           #statBlk := BLKMOV(SRCBLK := #identData, DSTBLK => #statWriteData);
           //Fill with data
           #statDat[4] := #statWriteData[#statWriteOffset];
           #statDat[5] := #statWriteData[1 + #statWriteOffset];
           #statDat[6] := #statWriteData[2 + #statWriteOffset];
           #statDat[7] := #statWriteData[3 + #statWriteOffset];
           #statDat[8] := #statWriteData[4 + #statWriteOffset];
           #statDat[9] := #statWriteData[5 + #statWriteOffset];
           #statDat[10] := #statWriteData[6 + #statWriteOffset];
           #statDat[11] := #statWriteData[7 + #statWriteOffset];
           #statDat[12] := #statWriteData[8 + #statWriteOffset];
           #statDat[13] := #statWriteData[9 + #statWriteOffset];
           #statDat[14] := #statWriteData[10 + #statWriteOffset];
           #statDat[15] := #statWriteData[11 + #statWriteOffset];
           #statDat[16] := #statWriteData[12 + #statWriteOffset];
           #statDat[17] := #statWriteData[13 + #statWriteOffset];
           #statDat[18] := #statWriteData[14 + #statWriteOffset];
           #statDat[19] := #statWriteData[15 + #statWriteOffset];
           #statDat[20] := #statWriteData[16 + #statWriteOffset];
           #statDat[21] := #statWriteData[17 + #statWriteOffset];
           #statDat[22] := #statWriteData[18 + #statWriteOffset];
           #statDat[23] := #statWriteData[19 + #statWriteOffset];
           #statDat[24] := #statWriteData[20 + #statWriteOffset];
           #statDat[25] := #statWriteData[21 + #statWriteOffset];
           #statDat[26] := #statWriteData[22 + #statWriteOffset];
           #statDat[27] := #statWriteData[23 + #statWriteOffset];
           #statDat[28] := #statWriteData[24 + #statWriteOffset];
           #statDat[29] := #statWriteData[25 + #statWriteOffset];
           #statDat[30] := #statWriteData[26 + #statWriteOffset];
           #statDat[31] := #statWriteData[27 + #statWriteOffset];

           //#statIOsizeNetto Bytes are reserved for every transfer
       END_IF;
       IF #statBlk = 0 THEN
           #statNState := #statTelegramState;                           //Telegram: Edit the read data
       END_IF;


       //-----------------------------------------------Telegram state----------------------------------------//
       //---------------------------------------------edit received data--------------------------------------//
       //-----------------------------------------------------------------------------------------------------//  

   1: //Telegram    
       IF #statLength > #statIOsizeNetto -1 THEN                 //Only when length of data > 0 can continue  
           IF #statStatusBits[6] THEN                            //IF RFID error has occured
               #tempStatusWord[1] := #statRecDat[1];          //error_RFID
               #tempStatusWord[0] := 16#0011;                          //Error identifier for RFID errors
               #status := #tempStatus;
               #statNState := #statErrorState;
           END_IF;

           //-------------------------- read command is ready------------------------------------------------//

           IF #statStatusBits[7] AND #statStatusBits[0] THEN
               IF #statRecDat[2] = #statAddrWrite[0] AND #statRecDat[3] = #statAddrWrite[1] THEN //received ADR must be ==sent ADR
                   IF #statBlk = 0 THEN
                       IF #statStatusBits[7] AND NOT #statStatusBits[6] THEN
                           #statLength := #statLength - #statIOsizeNetto;
                           //if len is not dividable with #statIOsizeNetto the adr offset has to be changed that the last (length < #statIOsizeNetto) command is done right
                           IF #statDiffToIOsizeNetto <> 0 AND #statLength < #statIOsizeNetto THEN
                               #statByteMove := #statIOsizeNetto - #statDiffToIOsizeNetto;
                           END_IF;
                           #statWriteOffset := #statWriteOffset + #statIOsizeNetto;                                   //offset must be changed
                           #statAddr := INT_TO_WORD(WORD_TO_INT(#statAddr) + #statIOsizeNetto);     //Change the ADR (#statIOsizeNetto Bytes)       
                           #statNState := #statWriteState;                      //Start a new read command
                       ELSE
                           #statNState := #statIdleState;
                       END_IF;
                   ELSE
                       #tempStatusWord[1] := INT_TO_WORD(#statBlk);                 //Error has to BLKMOV occured
                       #tempStatusWord[0] := 16#0001;                           //functions-Error identifier
                       #status := #tempStatus;
                       #statNState := #statErrorState;
                   END_IF;
               END_IF;
           END_IF;

       ELSE
           #statNState := #statIdleState;
           #statBusy := FALSE;
           #statDone := TRUE;
           #done := TRUE;
           #busy := FALSE;

           #statDat[0] := 16#0;                                          //Reset write command
           #InstSetIoPart(ID      := #hwID,
                          OFFSET  := #statAddrOffset,
                          LEN     := #statIOsize,
                          STATUS  => #statIoPartStatus,
                          ERROR   => #statIoPartError,
                          OUTPUTS := #statDat);

       END_IF;
       #InstSetIoPart(ID := #hwID,                              //read data from process image
                      OFFSET := #statAddrOffset,
                      LEN := #statIOsize,
                      STATUS => #statIoPartStatus,
                      ERROR => #statIoPartError,
                      OUTPUTS := #statDat);

       //------------------------------------------------------------------------------------------------------------//
       //-------------------------------------------------Error state------------------------------------------------//
       //---------------------------------------------error has occured----------------------------------------------//

   3://#Error_state
       #tempError := true;
       #error := #tempError;
       #statBusy := false;
       #statTImerIn := false;
       #statNState := #statIdleState;
       #statDone := false;

       #statDat[0] := 16#0;                                          //Reset write command
       #InstSetIoPart(ID      := #hwID,                              
                      OFFSET  := #statAddrOffset,
                      LEN     := #statIOsize,
                      STATUS  => #statIoPartStatus,
                      ERROR   => #statIoPartError,
                      OUTPUTS := #statDat);

   END_CASE;

   //------------------------------------------------------------------------------------------------------------//
   //-------------------------------------------------Timer------------------------------------------------------//
   //------------------------------------------------------------------------------------------------------------//

   #instTon(IN := #statTImerIn,
            PT := #statTimerPT);

   IF #instTon.Q THEN                      //error has occured. No tag on field during the 5 sec.
       #tempStatusWord[1] := 16#8101;                              //tag has left the field
       #tempStatusWord[0] := 16#0001;                              //identifier rfid errors
       #status:=#tempStatus;
       #statNState := #statErrorState;
   END_IF;
END_FUNCTION_BLOCK

FUNCTION_BLOCK "LIOLink_RF200_SwitchAntenna"   // FB4, SCL
TITLE = LRfidIOL_ANT
{ S7_Optimized_Access := 'FALSE' }
FAMILY : S7-300
VERSION : 3.1
// Set Antenna
// IO-Link V1.1
   VAR_INPUT
      execute : Bool;   // start process
      antennaState : Bool;   // set/reset antenna bit
      hwID : Word;   // Hardware identifier
      portAddr : Int;   // Start address of port
      "version" : Int := 11;
   END_VAR
   VAR_OUTPUT
      done : Bool;   // Ready
      busy : Bool;   // Block active
      error : Bool;   // Error has occured
      status : DWord;   // error status
      statusWord AT status : Array[0..1] of Word;
      presence : Bool;
   END_VAR
   VAR
      statExecuteReq : Bool;   // positive edge og execute
      statAntByte : Byte;   // Byte 0, Status byte
      statAntBit AT statAntByte : Array[0..7] of Bool;
      statNState : Int;   // current state
      statLastState : Int;   // last state
      statAntennaOn : Int := 1;   // On state
      statAntennaOff : Int := 2;   // OFF state
      statReadyState : Int := 3;
      statAnt : Array[0..31] of Byte;   // received buffer
      statAddrOffset : Int;   // step for FOR
      statSent : Array[0..31] of Byte;   // sent buffer
      statPresenceBit : Bool;
      statBusy : Bool;
      InstSetIoPart : SETIO_PART;
      statIoPartError : Bool;
      statIoPartStatus : DWord;
      InstGetIoPart : GETIO_PART;
      statIOsize : Int;
   END_VAR
   VAR_TEMP
      tempDone : Bool;
      tempError : Bool;
      tempStatus : DWord;
      tempStatus_W AT tempStatus : Array[0..1] of Word;
   END_VAR
   VAR CONSTANT
      IOL_V10 : Int := 8;
      IOL_V11 : Int := 32;
      VERSION_10 : Int := 10;   // Identifier IO-Link version 1.0
      VERSION_11 : Int := 11;   // Identifier IO-Link version 1.1
   END_VAR
BEGIN
   REGION BLOCK INFO HEADER
       //===============================================================================
       // Siemens / (c)Copyright 2020
       //-------------------------------------------------------------------------------
       // Title:            LIOLink_RF200_SwitchAntenna
       // Function:         Switches the antenna on/off of SIMATIC RF200 readers via IO-Link
       // Library:          LIOLink
       // Author:           Siemens Industry Online Support
       // Tested with:      CPU 317-2 PN/DP FW 3.2
       // Engineering:      TIA Portal V16
       // Restrictions:     --
       // Requirements:     --
       //-------------------------------------------------------------------------------
       // Change log table:
       // Version  | Date       | Expert in charge       | Changes applied
       //----------|------------|------------------------|------------------------------
       // 01.00.00 | 01.07.2013 | Online Support         | First release
       // 01.01.00 | 01.12.2016 | Online Support         | Upgrade to TIA Portal V14
       // 02.00.00 | 01.09.2017 | Online Support         | Upgrade to TIA Portal V14 SP1
       //                                                | Implementation of Programming styleguide
       //                                                | Added support for IO-Link V1.1 readers
       // 02.01.00 | 01.12.2017 | Online Support         | Bug fixes and performance improvements
       // 02.02.00 | 01.03.2020 | Online Support         | Upgrade to TIA Portal V16
       // 02.03.00 | 08.03.2020 | Online Support         | Added input "version" for IO-Link version
       //===============================================================================
   END_REGION

   IF #version = #VERSION_11 THEN                           //determine IO-Link reader version (1.0/1.1) to set offset
       #statIOsize := #IOL_V11;
   ELSE
       #statIOsize := #IOL_V10;
   END_IF;

   #statAddrOffset:=#portAddr;                              //start adress of port
   #InstGetIoPart(ID := #hwID,                              //read data from process image
                  OFFSET := #statAddrOffset,
                  LEN := #statIOsize,
                  STATUS => #statIoPartStatus,
                  ERROR => #statIoPartError,
                  INPUTS := #statAnt);

   #statAntByte:=#statAnt[0];                              //status byte
   #statPresenceBit := #statAntBit[5];                     //Presence bit. Transponder on field
   #presence := #statPresenceBit;
   #busy := #statBusy;

   //------------------------------------If error byte<>0--------------------------------------------------//
   //------------------------------------save the rfid error-----------------------------------------------//

   IF #statAnt[1]<>0 AND #statBusy THEN
     #statAntByte:=#statAnt[1];  
      #statusWord[1]:=BYTE_TO_WORD(#statAntByte);    //error_BLK
      #statusWord[0]:=16#0011;                    //identifier rfid errors
      #statBusy:=false;
      #done:=false;
      #error:=TRUE;
      #statNState:=0;
   END_IF;

   IF NOT #execute THEN
       #done := false;
       #error := false;
       #status := 0;
   END_IF;

   IF #execute AND #execute<>#statExecuteReq THEN //Positive Edge for antenna on
     #statLastState:=0;
     #statBusy:=TRUE;                              //Block active
     #done:=FALSE;                             //reset all output parameters
     #error:=FALSE;
     #status:=0;
     IF #antennaState THEN                          //if antenna then activate the ANTENNA_ON process
       #statNState:=#statAntennaOn;
     ELSIF NOT #antennaState THEN                   //if not antenna then activate the ANTENNA_OFF process 
       #statNState:=#statAntennaOff;
     END_IF;

   END_IF;
   #statExecuteReq:=#execute;


   //---------------------------------------Antenna on state-----------------------------------------------//
   //---------------------------------------Reset Antenna bit----------------------------------------------//

   CASE #statNState OF
       0:  //Idle
           ;
       1:  //Antenna_on
                                                        //Antenna on process
           #statAntBit[4] := false;                        //Reset Byte 0, bit 4
           #statSent[0] := 16#0;
           #statLastState := #statAntennaOn;
           #InstSetIoPart(ID := #hwID,                         //Write data into process image
                          OFFSET := #statAddrOffset,
                          LEN := #statIOsize,
                          STATUS => #statIoPartStatus,
                          ERROR => #statIoPartError,
                          OUTPUTS := #statSent);
           IF NOT #statIoPartError AND #statAnt[1] = 0 THEN
               #statNState := #statReadyState;
           ELSIF #statIoPartError THEN
               #tempError := true;
               #error := #tempError;                             //error has occured
               #statBusy := FALSE;
               #tempStatus_W[1] := DWORD_TO_WORD(#statIoPartStatus);//error_BLK
               #tempStatus_W[0] := 16#0001;                    //identifier block errors
           END_IF;
       2:
                                                      //Antenna off process
           #statAntBit[4] := true;                         //set Byte 0, bit 4
           #statSent[0] := 16#10;
           #statLastState := #statAntennaOff;
           #InstSetIoPart(ID := #hwID,                         //Write data into process image
                          OFFSET := #statAddrOffset,
                          LEN := #statIOsize,
                          STATUS => #statIoPartStatus,
                          ERROR => #statIoPartError,
                          OUTPUTS := #statSent);
           IF NOT #statIoPartError AND #statAnt[1] = 0 THEN
               IF #statAntByte = 16#10 THEN                    //if status_byte=16#10 then antenna off
                   #statNState := #statReadyState;
               END_IF;
           ELSIF #statIoPartError THEN
               #tempError := true;
               #error := #tempError;                              //Error has occured
               #statBusy := FALSE;
               #tempStatus_W[1] := DWORD_TO_WORD(#statIoPartStatus);//error_BLK
               #tempStatus_W[0] := 16#0001;                     //identifier block errors
           END_IF;
       3:
           #tempDone := true;
           #done := #tempDone;                           //Ready
           #statBusy := FALSE;
           #statNState := 0;
   END_CASE;
END_FUNCTION_BLOCK

// folder: LIOLink/S7-1200/1500/Base blocks

FUNCTION_BLOCK "LIOLink_Diagnose"   // FB3, SCL
TITLE = LIOLink_Diagnose
{ S7_Optimized_Access := 'TRUE' }
AUTHOR : SIOS
FAMILY : LIOLink
VERSION : 0.1
// LIOLink_Diagnose is used to read the diagnose of all the ports of any IO-Link-Master Product of Siemens.
   VAR_INPUT
      execute : Bool;   // Rising edge starts the execution of the action once
      hwID : HW_IO;   // Hardware identifier of IO-Link master module or first sub module
      cap : Int;   // Client Access Point (CAP) 0xB400 or 0x00E3 (227)
   END_VAR
   VAR_OUTPUT
      done : Bool;   // TRUE: FB processing successfully completed
      busy : Bool;   // TRUE: FB is active and new output values can be expected.
      error : Bool;   // FALSE: No error / TRUE: An error occurred during the execution of the FB.
      status : Word := 16#7000;   // 16#0000-16#7FFF: Status of the FB / 16#8000-16#FFFF: Error identification (see following table)
      diagnostics : "LIOLink_typeDiagnostics";   // Diagnostics information of FB
      events : "LIOLink_typeEvents";
   END_VAR
   VAR
      statExecuteOld : Bool;   // Previous value of input `execute` for edge detection
      statDone : Bool;   // Static value for output 'done'
      statBusy : Bool;   // Static value for output 'busy'
      statError : Bool;   // Static value for output 'error'
      statStatus : Word;   // Static value for output 'status'
      statSubFunctionStatus : DWord;   // Static value for output 'subFunctionStatus'.
      statFBState : DInt;   // State of the state machine
      statFBErrorState : DInt;   // State in the state machine of the block where the error occurred / Zustand in der Zustandsmaschine des Blocks, in dem der Fehler aufgetreten ist
      statHwID : HW_ANY;   // Static value for input 'HwID'
      statHwIDprevious : HW_IO;   // Static value for input 'hwID' from the previous execute / Statischer Wert für Eingang 'hwID'
      statEmptyDiagnostics : "LIOLink_typeDiagnostics";   // Empty diagnostics information (for initialization purposes only)
      instRdRec : RDREC;   // System function "read data record"
      instRdDiag : RDREC;   // System function "read data record"
      statDiagRecord : Array[0..#LAST_INDEX_DIAG_RECORD] of Byte;   // Data record of port diagnose
      statDiagRecordEco : "LIOLink_typeEvents";
      statCap : UInt;   // Static value for input 'cap'
      statRead : Array[0..231] of Byte;   // Data record, Output of RDREC
      statIndexDiag : UInt;   // Static value for index of data record of port diagnose
      statPortNumber : Int := 8;   // Number of Ports of IO-Link-Master
      statPortEco : UInt := 1;   // Static value for a port counter of EcoPN
   END_VAR
   VAR_TEMP
      tempExecute : Bool;   // Temporary value for input 'execute'
      tempHwID : HW_IO;   // Temporary value for input 'hwID'
      tempCap : Int;   // Temporary value for input 'cap'
      tempPortNumber : Int;   // Temporary value for port number
      tempEventNumber : Int;   // Temporary value for event number
      tempIndexDiagRec : Int;   // Temporary value for index of data record (array) of diagnose
   END_VAR
   VAR CONSTANT
      INDEX_CAP_IOLINK : Word := 16#B000;   // Index of the data record for IOLM_Info. Only IO-Link-Masters with CAP=16#B000 support this call.
      INDEX_DIAG_OTHER : Word := 16#00E5;   // Index for port status based on Siemens Standard (old): 229 => reads status of all ports
      INDEX_DIAG_ECO : Word := 16#B200;   // Index for port status based on IO-Link-Standard: 16#B20n, n:Port number => reads port status of only one port
      CAP_LEGACY : Word := 16#00E3;   // Siemens (old) Standard CAP: 227
      CAP_STANDARD : Word := 16#B400;   // IO-Link Standard CAP: 16#B400
      STATUS_EXECUTION_FINISHED_NO_ERROR : Word := 16#0000;   // Processing finished without error
      STATUS_NO_CALL : Word := 16#7000;   // No current processing request / no order in process
      STATUS_FIRST_CALL : Word := 16#7001;   // First call after new incoming job request (rising edge at 'execute')
      STATUS_SUBSEQUENT_CALL : Word := 16#7002;   // Subfunction call in progress without further detailing
      STATUS_MASK : DWord := 16#00FF_FF00;   // Mask to filter error codes
      STATUS_RESOURCE_BUSY : DWord := 16#0080_C200;   // Status from WRREC/RDREC: Resource is busy
      ERR_UNDEFINED_STATE : Word := 16#8600;   // Error in function due to an undefined state in the state machine
      ERR_RDREC : Word := 16#8602;   // Error: RDREC encountered an error, see "diagnostics"
      FB_STATE_NO_PROCESSING : DInt := 0;   // FB state: No processing
      FB_STATE_READ_CAP : DInt := 1;   // FB state: Read CAP
      FB_STATE_READ_DIAG : DInt := 2;   // FB state: Read diagnose
      MIN_PORT : Int := 1;   // Minimum number of ports
      MAX_PORT : Int := 8;   // Maximum number of ports
      MIN_EVENTS : Int;   // Minimum number of events
      MAX_EVENTS : Int := 4;   // Maximum number of events
      MASTER_PORT_STATUS_V2 : Byte := 16#02;   // Master port status version 2
      MASTER_PORT_STATUS_V3 : Byte := 16#03;   // Master port status version 3
      MASTER_PORT_STATUS_V4 : Byte := 16#04;   // Master port status version 4
      START_INDEX_MASTER_PORT_STATUS_V2 : Int := 28;   // Start index of relevant data in the case of port status version 2
      START_INDEX_MASTER_PORT_STATUS_V3 : Int := 34;   // Start index of relevant data in the case of port status version 3
      START_INDEX_MASTER_PORT_STATUS_V4 : Int := 42;   // Start index of relevant data in the case of port status version 4
      START_INDEX_MASTER_PORT_STATUS_STANDARD : Int := 18;   // Start index of relevant data in case of a IO-Link Standard data record for port status
      START_INDEX_DIAG_RECORD : Int := 0;   // Start index of diagnose record array
      LAST_INDEX_DIAG_RECORD : Int := 231;   // Last index of diagnose record array
      RESET_WORD : Word := 16#0000;   // Reset event codes
      RESET_BYTE : Byte := 16#00;   // Reset byte for statDiagRecord
      STATUS_RDREC_VALID : Byte := 16#00;   // Status Code of RDREC in cased of no error occurs
      BITMASK_ERR_RDREC_B3 : Byte := 16#DE;   // Status Code of RDREC in case of an error when reading a data record
      BITMASK_ERR_RDREC_B2 : Byte := 16#80;   // Status Code of RDREC in case of an error when reading a data record - Error according to IEC 61158-6
      BITMASK_ERR_RDREC_B1 : Byte := 16#B0;   // Status Code of RDREC in case of an error when reading a data record - invalid index (cap)
   END_VAR
BEGIN
   REGION BLOCK INFO HEADER
       //===============================================================================
       // Siemens / (c)Copyright 2023
       //-------------------------------------------------------------------------------
       // Title:            LIOLink_Diagnosis
       // Function:         Reads diagnose of ports of IO-Link-Masters in IO-Link Standard
       // Library:          LIOLink
       // Author:           SUP SPH
       // Tested with:      CPU 1511F-1 PN FW 2.8
       // Engineering:      TIA Portal V16
       // Restrictions:     S7-1200/1500
       // Requirements:     --
       //-------------------------------------------------------------------------------
       // Change log table:
       // Version  | Date       | Expert in charge       | Changes applied
       //----------|------------|------------------------|------------------------------
       // 01.00.00 | 28.02.2023 | SUP SPH                | First release for TIA Portal V16
       // 
       //===============================================================================
   END_REGION


   REGION TRIGGERING
       #tempExecute := #execute; // Work with temporary value / create process image

       IF (#tempExecute = TRUE) AND (#statExecuteOld = FALSE) // Check if FB is triggered
           // FB shall finish current job before new job can be started with rising edge of execute
           AND (#statStatus = #STATUS_NO_CALL)
       THEN
           REGION Initialize data
               // First call; initialize FB
               #statDone := FALSE;
               #statBusy := TRUE;
               #statError := FALSE;
               #statStatus := #STATUS_FIRST_CALL;
               #statSubFunctionStatus := #STATUS_EXECUTION_FINISHED_NO_ERROR;
               #statFBErrorState := 0;
               #diagnostics := #statEmptyDiagnostics;
               //save the hwID from the previous execute
               #statHwIDprevious := #statHwID;

               //reset static variables of Diagnose Records
               FOR #tempPortNumber := #MIN_PORT TO #MAX_PORT DO
                   FOR #tempEventNumber := #MIN_EVENTS TO #MAX_EVENTS DO
                       #statDiagRecordEco."port"[#tempPortNumber].event[#tempEventNumber].eventQualifier.instance := #RESET_BYTE;
                       #statDiagRecordEco."port"[#tempPortNumber].event[#tempEventNumber].eventQualifier.source := FALSE;
                       #statDiagRecordEco."port"[#tempPortNumber].event[#tempEventNumber].eventQualifier.type := #RESET_BYTE;
                       #statDiagRecordEco."port"[#tempPortNumber].event[#tempEventNumber].eventQualifier.mode := #RESET_BYTE;
                       #statDiagRecordEco."port"[#tempPortNumber].event[#tempEventNumber].eventCode := #RESET_WORD;
                   END_FOR;
               END_FOR;
               FOR #tempIndexDiagRec := #START_INDEX_DIAG_RECORD TO #LAST_INDEX_DIAG_RECORD DO
                   #statDiagRecord[#tempIndexDiagRec] := #RESET_BYTE;
               END_FOR;
           END_REGION

           REGION Save inputs
               //save input parameters
               #tempHwID := #hwID;
               #tempCap := #cap;
           END_REGION

           REGION Check parameters
               IF #statStatus = #STATUS_FIRST_CALL THEN // Parameters OK
                   IF #tempCap <> 0 THEN   //check if cap is predefined, or given by the user
                       #statCap := INT_TO_UINT(#tempCap);
                       #statFBState := #FB_STATE_READ_DIAG;
                   ELSIF (#statCap <> WORD_TO_UINT(#CAP_STANDARD) AND #statCap <> WORD_TO_UINT(#CAP_LEGACY)) OR (#statHwIDprevious <> #tempHwID) THEN
                       #statFBState := #FB_STATE_READ_CAP;
                   ELSE //CAP already known
                       #statFBState := #FB_STATE_READ_DIAG;
                   END_IF;
               END_IF;
               //save current hwID
               #statHwID := #tempHwID;
           END_REGION

       ELSIF (#statStatus = #STATUS_FIRST_CALL) THEN
           #statStatus := #STATUS_SUBSEQUENT_CALL;
       ELSIF (#statFBState=#FB_STATE_NO_PROCESSING) THEN
           #statStatus := #STATUS_NO_CALL;
           #statDone := FALSE;
           #statBusy := FALSE;
           #statError := FALSE;

           #instRdDiag(REQ := FALSE,
                       RECORD := #statDiagRecord);

           #instRdRec(REQ := FALSE,
                      RECORD := #statRead);
       END_IF;

       // Edge detection 'execute' input
       #statExecuteOld := #tempExecute;
   END_REGION TRIGGERING

   REGION STATE_MACHINE
       CASE #statFBState OF // State machine of FB
           #FB_STATE_NO_PROCESSING: // No processing active (Note: this state must always be present and left empty)
               REGION No processing
                   ;
               END_REGION

           #FB_STATE_READ_CAP:
               REGION Read CAP
                   // To find out CAP of IO-Link Master, data record with Index 16#B000 is read. If this reading was successful
                   // then CAP is 16#B400 (based on IO-Link Standard). If the reading was not successful and the status of RDREC
                   // is 16#DE80_B0xx, then CAP is 16#00E3 (227, based on Siemens Old Standard for IO-Link Masters).

                   #instRdRec(RECORD := #statRead);

                   IF (#instRdRec.BUSY = FALSE) THEN
                       IF (#instRdRec.VALID = FALSE) AND (#instRdRec.ERROR = FALSE) THEN
                           IF #instRdRec.REQ = FALSE THEN
                               // call read record with Index 16#B000
                               #instRdRec.REQ := TRUE;
                               #instRdRec.ID := #statHwID;
                               #instRdRec.INDEX := WORD_TO_UINT(#INDEX_CAP_IOLINK);
                               #instRdRec.MLEN := 0;
                               #statFBState := #FB_STATE_READ_CAP;
                           END_IF;
                       ELSIF #instRdRec.VALID = TRUE THEN
                           #instRdRec.REQ := FALSE;
                           // if status of RDREC is valid then CAP is 16#B400 (CAP_STANDARD)
                           IF #instRdRec.STATUS.%B3 = #STATUS_RDREC_VALID THEN
                               #statCap := WORD_TO_UINT(#CAP_STANDARD);
                               #statPortNumber := BYTE_TO_INT(#statRead[11]); //read number of ports of IO-Link-Master
                               #statPortEco := 1;
                               #statIndexDiag := WORD_TO_UINT(#INDEX_DIAG_ECO) + #statPortEco; //Data Record with the status of each port: 0xB20n, n - Port number
                           END_IF;
                           #statFBState := #FB_STATE_READ_DIAG;
                       ELSE
                           // if RDREC is in error state and Status is 16#DE80_B0xx then CAP is 227 (CAP_Legacy)
                           IF (#instRdRec.STATUS.%B3 = #BITMASK_ERR_RDREC_B3) AND (#instRdRec.STATUS.%B2 = #BITMASK_ERR_RDREC_B2) AND (#instRdRec.STATUS.%B1 = #BITMASK_ERR_RDREC_B1) THEN
                               #statCap := WORD_TO_UINT(#CAP_LEGACY);
                               #statIndexDiag := WORD_TO_UINT(#INDEX_DIAG_OTHER);
                               #statFBState := #FB_STATE_READ_DIAG;
                           ELSE
                               #statDone := FALSE;
                               #statBusy := FALSE;
                               #statError := TRUE;
                               #statStatus := #ERR_RDREC;
                               #statCap := 0; //clear CAP if an error occurs
                               #statIndexDiag := 0;
                               #statSubFunctionStatus := #instRdRec.STATUS;
                               #statFBErrorState := #statFBState;
                               #statFBState := #FB_STATE_NO_PROCESSING;
                           END_IF;
                       END_IF;
                   ELSE
                       #instRdRec.REQ := FALSE;
                   END_IF;

                   #instRdRec(RECORD := #statRead);
               END_REGION

           #FB_STATE_READ_DIAG:
               REGION Read Diagnosis

                   REGION read diagnosis in case of Siemens-Version //statIndex 229
                       //diagnose of all ports is read with only one call
                       IF #statIndexDiag = WORD_TO_UINT(#INDEX_DIAG_OTHER) THEN
                           #instRdDiag(RECORD := #statDiagRecord);
                           IF (#instRdDiag.BUSY = FALSE) THEN
                               IF (#instRdDiag.VALID = FALSE) AND (#instRdDiag.ERROR = FALSE) THEN
                                   IF #instRdDiag.REQ = FALSE THEN
                                       #instRdDiag.REQ := TRUE;
                                       #instRdDiag.ID := #statHwID;
                                       #instRdDiag.INDEX := #statIndexDiag;
                                       #instRdDiag.MLEN := 0;
                                   END_IF;
                               ELSE
                                   #instRdDiag.REQ := FALSE;
                                   IF #instRdDiag.VALID = TRUE THEN  //Diagnose valid, statDone is true
                                       #statStatus := #STATUS_EXECUTION_FINISHED_NO_ERROR;
                                       #statFBState := #FB_STATE_NO_PROCESSING;
                                       #statDone := TRUE;
                                       #statBusy := FALSE;
                                       #statError := FALSE;
                                   ELSE
                                       IF (#instRdDiag.STATUS AND #STATUS_MASK) <> #STATUS_RESOURCE_BUSY THEN  //Error occured
                                           #statDone := FALSE;
                                           #statBusy := FALSE;
                                           #statError := TRUE;
                                           #statStatus := #ERR_RDREC;
                                           #statCap := 0;
                                           #statIndexDiag := 0;
                                           #statSubFunctionStatus := #instRdDiag.STATUS;
                                           #statFBErrorState := #statFBState;
                                           #statFBState := #FB_STATE_NO_PROCESSING;
                                       END_IF;
                                   END_IF;
                               END_IF;
                           ELSE
                               #instRdDiag.REQ := FALSE;
                           END_IF;
                           #instRdDiag(RECORD := #statDiagRecord);
                       END_IF;
                   END_REGION

                   REGION read diagnosis in case of Standard-Version // Index 0xB20n, n - Port number
                       IF #statIndexDiag = (WORD_TO_UINT(#INDEX_DIAG_ECO) + #statPortEco) THEN
                           //one call for each port diagnose, statPortEco starting from 1 to maximum number of ports
                           IF #statPortEco < (#statPortNumber + 1) THEN
                               #instRdDiag(RECORD := #statDiagRecord);
                               IF (#instRdDiag.BUSY = FALSE) THEN
                                   IF (#instRdDiag.VALID = FALSE) AND (#instRdDiag.ERROR = FALSE) THEN
                                       IF #instRdDiag.REQ = FALSE THEN
                                           #instRdDiag.REQ := TRUE;
                                           #instRdDiag.ID := #statHwID;
                                           #instRdDiag.INDEX := #statIndexDiag;
                                           #instRdDiag.MLEN := 0;
                                       END_IF;
                                   ELSE
                                       #instRdDiag.REQ := FALSE;
                                       IF #instRdDiag.VALID = TRUE THEN  //Diagnose of port is valid
                                           #tempIndexDiagRec := #START_INDEX_MASTER_PORT_STATUS_STANDARD; //starting index of data record, where events are recorded
                                           //for each port, the 5 last-events are saved in output
                                           FOR #tempEventNumber := #MIN_EVENTS TO #MAX_EVENTS DO
                                               #statDiagRecordEco."port"[#statPortEco].event[#tempEventNumber].eventQualifier.instance.%X0 := #statDiagRecord[#tempIndexDiagRec].%X0;
                                               #statDiagRecordEco."port"[#statPortEco].event[#tempEventNumber].eventQualifier.instance.%X1 := #statDiagRecord[#tempIndexDiagRec].%X1;
                                               #statDiagRecordEco."port"[#statPortEco].event[#tempEventNumber].eventQualifier.instance.%X2 := #statDiagRecord[#tempIndexDiagRec].%X2;
                                               #statDiagRecordEco."port"[#statPortEco].event[#tempEventNumber].eventQualifier.source := #statDiagRecord[#tempIndexDiagRec].%X3;
                                               #statDiagRecordEco."port"[#statPortEco].event[#tempEventNumber].eventQualifier.type.%X0 := #statDiagRecord[#tempIndexDiagRec].%X4;
                                               #statDiagRecordEco."port"[#statPortEco].event[#tempEventNumber].eventQualifier.type.%X1 := #statDiagRecord[#tempIndexDiagRec].%X5;
                                               #statDiagRecordEco."port"[#statPortEco].event[#tempEventNumber].eventQualifier.mode.%X0 := #statDiagRecord[#tempIndexDiagRec].%X6;
                                               #statDiagRecordEco."port"[#statPortEco].event[#tempEventNumber].eventQualifier.mode.%X1 := #statDiagRecord[#tempIndexDiagRec].%X7;
                                               #statDiagRecordEco."port"[#statPortEco].event[#tempEventNumber].eventCode.%B1 := #statDiagRecord[#tempIndexDiagRec + 1];
                                               #statDiagRecordEco."port"[#statPortEco].event[#tempEventNumber].eventCode.%B0 := #statDiagRecord[#tempIndexDiagRec + 2];
                                               #tempIndexDiagRec := #tempIndexDiagRec + 3; //3-bytes for each event => 2 bytes for event code + 1 byte for event type
                                           END_FOR;
                                           #statPortEco := #statPortEco + 1; //port number is updated => next port
                                           #statIndexDiag := WORD_TO_UINT(#INDEX_DIAG_ECO) + #statPortEco; //change index for the next port diagnose
                                       ELSE
                                           IF (#instRdDiag.STATUS AND #STATUS_MASK) <> #STATUS_RESOURCE_BUSY THEN  //Error occured
                                               #statDone := FALSE;
                                               #statBusy := FALSE;
                                               #statError := TRUE;
                                               #statStatus := #ERR_RDREC;
                                               #statCap := 0;
                                               #statIndexDiag := 0;
                                               #statSubFunctionStatus := #instRdDiag.STATUS;
                                               #statFBErrorState := #statFBState;
                                               #statFBState := #FB_STATE_NO_PROCESSING;
                                               #statPortEco := 0;
                                           END_IF;
                                       END_IF;
                                   END_IF;
                               ELSE
                                   #instRdDiag.REQ := FALSE;
                               END_IF;
                               #instRdDiag(RECORD := #statDiagRecord);
                           ELSE
                               //diagnose of all ports was successfully read
                               #statPortEco := 1;
                               #statIndexDiag := WORD_TO_UINT(#INDEX_DIAG_ECO) + #statPortEco;
                               #statStatus := #STATUS_EXECUTION_FINISHED_NO_ERROR;
                               #statFBState := #FB_STATE_NO_PROCESSING;
                               #statDone := TRUE;
                               #statBusy := FALSE;
                               #statError := FALSE;
                           END_IF;
                       END_IF;
                   END_REGION


               END_REGION

           ELSE // Undefined state in state machine reached
               #statDone := FALSE;
               #statBusy := FALSE;
               #statError := TRUE;
               #statStatus := #ERR_UNDEFINED_STATE;
       END_CASE;
   END_REGION STATE_MACHINE

   REGION OUTPUTS
       // Write outputs

       // Fill event codes in case of new received diagnosis data
       IF #statDone = TRUE THEN
           IF #statIndexDiag = WORD_TO_UINT(#INDEX_DIAG_OTHER) THEN
               //Diagnosis record in case of Siemens Old Standard
               REGION EVENTCODES_SIEMENS_VERSION
                   //The master post status record has 3 versions (1,2,3-Version). For each post status record there is a different offset, from where the diagnose data can be found.
                   //The master port status version is found in Byte 0 of each port status data record e.g. statDiagRecord[0].
                   //Therefore based on the master port status version, the start index of diagnose data is found.
                   IF #statDiagRecord[0] = #MASTER_PORT_STATUS_V2 THEN
                       #tempIndexDiagRec := #START_INDEX_MASTER_PORT_STATUS_V2;
                   ELSIF #statDiagRecord[0] = #MASTER_PORT_STATUS_V3 THEN
                       #tempIndexDiagRec := #START_INDEX_MASTER_PORT_STATUS_V3;
                   ELSIF #statDiagRecord[0] = #MASTER_PORT_STATUS_V4 THEN
                       #tempIndexDiagRec := #START_INDEX_MASTER_PORT_STATUS_V4;
                   END_IF;

                   IF (#statDiagRecord[0] = #MASTER_PORT_STATUS_V2) OR (#statDiagRecord[0] = #MASTER_PORT_STATUS_V3) OR (#statDiagRecord[0] = #MASTER_PORT_STATUS_V4) THEN
                       FOR #tempPortNumber := #MIN_PORT TO #MAX_PORT DO
                           FOR #tempEventNumber := #MIN_EVENTS TO #MAX_EVENTS DO
                               #events."port"[#tempPortNumber].event[#tempEventNumber].eventQualifier.instance.%X0 := #statDiagRecord[#tempIndexDiagRec].%X0;
                               #events."port"[#tempPortNumber].event[#tempEventNumber].eventQualifier.instance.%X1 := #statDiagRecord[#tempIndexDiagRec].%X1;
                               #events."port"[#tempPortNumber].event[#tempEventNumber].eventQualifier.instance.%X2 := #statDiagRecord[#tempIndexDiagRec].%X2;
                               #events."port"[#tempPortNumber].event[#tempEventNumber].eventQualifier.source := #statDiagRecord[#tempIndexDiagRec].%X3;
                               #events."port"[#tempPortNumber].event[#tempEventNumber].eventQualifier.type.%X0 := #statDiagRecord[#tempIndexDiagRec].%X4;
                               #events."port"[#tempPortNumber].event[#tempEventNumber].eventQualifier.type.%X1 := #statDiagRecord[#tempIndexDiagRec].%X5;
                               #events."port"[#tempPortNumber].event[#tempEventNumber].eventQualifier.mode.%X0 := #statDiagRecord[#tempIndexDiagRec].%X6;
                               #events."port"[#tempPortNumber].event[#tempEventNumber].eventQualifier.mode.%X1 := #statDiagRecord[#tempIndexDiagRec].%X7;
                               #events."port"[#tempPortNumber].event[#tempEventNumber].eventCode.%B1 := #statDiagRecord[#tempIndexDiagRec + 1];
                               #events."port"[#tempPortNumber].event[#tempEventNumber].eventCode.%B0 := #statDiagRecord[#tempIndexDiagRec + 2];
                               #tempIndexDiagRec := #tempIndexDiagRec + 3; //3-bits for each event, 2 bits for eventcode + 1 bit for event type
                           END_FOR;
                           #tempIndexDiagRec := #tempIndexDiagRec + 4; //4 bits reserved for other purposes between Port Diagnoses
                       END_FOR;
                   END_IF;
               END_REGION
               //Diagnosis record in case of IO-Link-Standard
           ELSIF #statIndexDiag = (WORD_TO_UINT(#INDEX_DIAG_ECO) + #statPortEco) THEN
               REGION EVENTCODES_STANDARD_VERSION
                   #events := #statDiagRecordEco;
               END_REGION
           END_IF;
       ELSIF #statError = TRUE THEN  //Error occurred
           #diagnostics.status := #statStatus;
           #diagnostics.subfunctionStatus := #statSubFunctionStatus;
           #diagnostics.stateNumber := #statFBErrorState;
       END_IF;

       // Write static function block status values to outputs
       #done := #statDone;
       #busy := #statBusy;
       #error := #statError;
       #status := #statStatus;

   END_REGION OUTPUTS
END_FUNCTION_BLOCK

FUNCTION_BLOCK "LIOLink_Device"   // FB50004, SCL
TITLE = LIOLink_Device / LIOLINK_DEVICE
{ S7_Optimized_Access := 'TRUE' }
AUTHOR : SIOS
FAMILY : LIOLink
VERSION : 4.0
// Acyclically reads or writes data records from and to IO-Link devices / Funktionsbaustein zum Lesen und Schreiben von azyklischen Daten auf Geräten mit IO-Link, die auf SIMATIC S7-Steuerungen verwendet werden. (früher IO_LINK_CALL)
   VAR_INPUT
      execute : Bool;   // Request to execute function / Anforderung zum Ausführen der Funktion
      hwID : HW_IO;   // Hardware identifier of IO-Link master module or first sub module / Hardware-Kennung des IO-Link-Mastermoduls (Submodul für ET 200eco PN)
      cap : Int;   // Client Access Point (CAP) 0xB400 or 0x00E3 (227) / Client Access Point (CAP); 0xB400 für ET 200eco PN, CM 8x IO-Link, sonst 0xE003 (227)
      readWrite : Bool;   // FALSE: read-mode, TRUE: write-mode / FALSE: lesen, TRUE: schreiben
      port : Int;   // Port on IO-Link master module / Port am IO-Link-Master-Modul
      index : Int;   // Address parameter index (IO-Link device); 0..32767: IOL-D; 65535: port functions / Adressparameterindex (IO-Link Device); 0..32767: IOL-D; 65535: Portfunktionen
      subindex : Int;   // Address parameter subindex (IO-Link device); 0: full record; 1-255: single parameter / Adressparameter Subindex (IO-Link Device); 0: vollständige Aufzeichnung; 1-255: Einzelparameter
      writeLen : Int;   // Length of writing data (net data); 1..232 / Länge der Schreibdaten (Nettodaten); 1..232
      timeout : Time := T#20S;   // Time after which the request is aborted / Zeit, nach der die Anfrage abgebrochen wird
      pollingPeriod : Time := T#100MS;   // Time period of polling
   END_VAR
   VAR_OUTPUT
      done : Bool;   // TRUE: FB processing successfully completed / TRUE: FB-Bearbeitung erfolgreich abgeschlossen
      busy : Bool;   // TRUE: FB is active and new output values can be expected. / TRUE: FB ist aktiv und neue Ausgangswerte sind zu erwarten.
      error : Bool;   // FALSE: No error / TRUE: An error occurred during the execution of the FB. / FALSE: Kein Fehler / TRUE: Bei der Ausführung des FB ist ein Fehler aufgetreten.
      status : Word := 16#7000;   // 16#0000-16#7FFF: Status of the FB / 16#8000-16#FFFF: Error identification (see following table) / 16#0000-16#7FFF: Status des FB / 16#8000-16#FFFF: Fehleridentifikation (siehe folgende Tabelle)
      diagnostics : "LIOLink_typeDiagnostics";   // Diagnostics information of FB / Diagnoseinformationen der FB
      readLen : Int;   // Length of read data record (number of bytes) / Länge des gelesenen Datensatzes (Anzahl Bytes)
   END_VAR
   VAR_IN_OUT
      record : Array[*] of Byte;   // Data area for reading/writing data (max. 232 byte) / Datenbereich zum Lesen/Schreiben von Daten (max. 232 Byte)
   END_VAR
   VAR
      statExecuteOld : Bool;   // Old value of 'execute' input for edge detection / Alter Wert des 'Execute'-Eingangs für Flankenerkennung
      statDone : Bool;   // Static value for output 'done' / Statischer Wert für Ausgang 'done'
      statBusy : Bool;   // Static value for output 'busy' / Statischer Wert für Ausgang 'besetzt'
      statError : Bool;   // Static value for output 'error' / Statischer Wert für Ausgang 'error'
      statStatus : Word := 16#7000;   // Static value for output 'status' / Statischer Wert für Ausgang 'Status'
      statPollingPeriod : Time := T#100MS;   // Static value for input 'pollingPeriod'
      statHwID : HW_IO;   // Static value for input 'hwID' / Statischer Wert für Eingang 'hwID'
      statHwIDprevious : HW_IO;   // Static value for input 'hwID' from the previous execute / Statischer Wert für Eingang 'hwID'
      statReadWrite : Bool;   // Static value for input 'readWrite' / Stativwert für Eingabe 'readWrite'
      statCap : UInt;   // Static value for input 'cap' / Statischer Wert für Eingabe 'cap'
      statTimeout : Time;   // Static value for input 'timeout' / Statischer Wert für Eingang 'timeout'
      statLen : UInt;   // Length of data to be written to device / Länge der Daten, die auf das Gerät geschrieben werden sollen
      statSubfunctionStatus : DWord;   // Status of WRREC/RDREC or error code from IO-Link Master (%W1: IO-Link Master error, %W0: ISDU error) / Status von WRREC/RDREC oder Fehlercode vom IO-Link-Master (%W1: IO-Link-Master-Fehler, %W0: ISDU-Fehler)
      statFBErrorState : DInt;   // State in the state machine of the block where the error occurred / Zustand in der Zustandsmaschine des Blocks, in dem der Fehler aufgetreten ist
      statFBState : DInt := 0;   // State in the state machine of the FB / Zustand in der Zustandsmaschine der FB
      statEmptyDiagnostics : "LIOLink_typeDiagnostics";   // Empty diagnostics information (for initialization purposes only) / Leere Diagnoseinformationen (nur für Initialisierungszwecke)
      instRdRec : RDREC;   // System function "read data record" / Systemfunktion "Datensatz lesen"
      instWrRec : WRREC;   // System function "write data record" / Systemfunktion "Datensatz schreiben"
      instPoll : TP_TIME;   // poll rate read data record / Abfragerate Datensatz lesen
      instMonitor : TON_TIME;   // request monitoring time / Überwachungszeit anfordern
      statRead : Struct   // data area for reading data / Datenbereich zum Lesen von Daten
         header : Struct   // Header
            call : Struct   // header for read/write data record / Header für Datensatz lesen/schreiben
               extFunctionNum : Byte := 16#08;   // extended function number (fix coded 08h) / erweiterte Funktionsnummer (fix codiert 08h)
               port : Byte;   // variable port (user interface) 0...255 / variabler Port (Benutzeroberfläche) 0...255
               fiIndex : Word := 16#FE4A;   // FI index (fix coded 65098) / FI-Index (fix codiert 65098)
            END_STRUCT;
            iolHeader : Struct   // header for IO-Link / Header für IO-Link
               control : Byte;   // RD_WR = 0 = read = Control:=0x03 / / RD_WR = 1 = write = Control:=0x02 / RD_WR = 0 = lesen = Steuerung:=0x03 / / RD_WR = 1 = schreiben = Steuerung:=0x02
               indexHighByte : Byte;   // index of data record 0…32767 (high byte) / Index des Datensatzes 0…32767 (High Byte)
               indexLowByte : Byte;   // index of data record 0…32767 (low byte) / Index des Datensatzes 0…32767 (Low Byte)
               subindex : Byte;   // subindex for data record 0...255 / Subindex für Datensatz 0...255
            END_STRUCT;
         END_STRUCT;
         data : Array[0..231] of Byte;   // Data
      END_STRUCT;
      statWrite : Struct   // data area for writing data / Datenbereich zum Schreiben von Daten
         header : Struct   // Header
            call : Struct   // header for read/write data record / Header für Datensatz lesen/schreiben
               extFunctionNum : Byte := 16#08;   // extended function number (fix coded 08h) / erweiterte Funktionsnummer (fix codiert 08h)
               port : Byte;   // variable port (user interface) 0...255 / variabler Port (Benutzeroberfläche) 0...255
               fiIndex : Word := 16#FE4A;   // FI index (fix coded 65098) / FI-Index (fix codiert 65098)
            END_STRUCT;
            iolHeader : Struct   // header für IO-Link / Header für IO-Link
               control : Byte;   // RD_WR = 0 = read = Control:=0x03 / / RD_WR = 1 = write = Control:=0x02 / RD_WR = 0 = lesen = Steuerung:=0x03 / / RD_WR = 1 = schreiben = Steuerung:=0x02
               indexHighByte : Byte;   // index of data record 0…32767 (high byte) / Index des Datensatzes 0…32767 (High Byte)
               indexLowByte : Byte;   // index of data record 0…32767 (low byte) / Index des Datensatzes 0…32767 (Low Byte)
               subindex : Byte;   // subindex for data record 0...255 / Subindex für Datensatz 0...255
            END_STRUCT;
         END_STRUCT;
         data : Array[0..231] of Byte;   // Data
      END_STRUCT;
   END_VAR
   VAR_TEMP
      tempExecute : Bool;   // Temporary value for input 'execute' / Temporärer Wert für Eingabe 'execute'
      tempHwID : HW_IO;   // Temporary value for input 'hwID'
      tempPort : Int;   // Temporary value for input 'port'
      tempIndex : Int;   // Temporary value for input 'index'
      tempSubindex : Int;   // Temporary value for input 'subindex'
      tempIndexCounter : DInt;   // run tag for counting loops / Run-Tag für Zählschleifen
   END_VAR
   VAR CONSTANT
      MODE_READ : Bool := FALSE;   // Mode to read data / Modus zum Lesen von Daten
      MODE_WRITE : Bool := TRUE;   // Mode to write data / Modus zum Schreiben von Daten
      MAX_PORT : USInt := 63;   // Max. possible port / max. möglichen Hafen
      MAX_INDEX : UInt := 32767;   // Max. possible index / max. möglicher Index
      INDEX_PORT_FUNC : UInt := 65535;   // Index to address port functions / Index zum Adressieren von Portfunktionen
      MAX_SUBINDEX : USInt := 255;   // Max. possible subindex / max. möglicher Subindex
      MAX_DATA : USInt := 232;   // Max. size of data to be transferred / max. Größe der zu übertragenden Daten
      UPPER_LIMIT : DInt := 231;   // Upper limit of data to be transferred / Obergrenze der zu übertragenden Daten
      FB_STATE_NO_PROCESSING : DInt := 0;   // FB state: No processing / FB-Zustand: Keine Verarbeitung
      FB_STATE_WRITE : DInt := 1;   // FB state: Write data record / Datensatz schreiben
      FB_STATE_POLL : DInt := 2;   // FB state: Wait and poll for response / warten und auf Antwort abfragen
      FB_STATE_READ_CAP : DInt := 3;   // FB state: Read cap / CAP lesen
      IOL_HEADER : UInt := 65098;   // Header IO-Link / Kopfzeile IO-Link
      LEN_HEADER : USInt := 8;   // Length of header / Länge des Headers
      CONTROL_WRITE : Byte := 16#02;   // Write data record / Datensatz schreiben
      CONTROL_READ : Byte := 16#03;   // Read data record / Datensatz lesen
      STATUS_EXECUTION_FINISHED : Word := 16#0000;   // Execution finished without errors / Ausführung ohne Fehler beendet
      STATUS_NO_CALL : Word := 16#7000;   // No job being currently processed / Derzeit wird kein Auftrag bearbeitet
      STATUS_FIRST_CALL : Word := 16#7001;   // First call after incoming new job (rising edge 'execute') / Erster Aufruf nach eingehendem neuen Auftrag (steigende Flanke 'execute')
      STATUS_SUBSEQUENT_CALL : Word := 16#7002;   // Subsequent call during active processing without further details / Nachfolgender Aufruf während aktiver Bearbeitung ohne weitere Angaben
      SUB_STATUS_NO_ERROR : Word := 16#0000;   // No error occured in subfunction call / Fehler: falscher Port
      ERR_WRONG_PORT : Word := 16#8201;   // Error: wrong port / Fehler: falscher Index
      ERR_WRONG_INDEX : Word := 16#8202;   // Error: wrong index / Fehler: falscher Subindex
      ERR_WRONG_SUBINDEX : Word := 16#8203;   // Error: wrong subindex / Fehler: falsche Länge für Datensatz schreiben
      ERR_WRONG_LENGTH : Word := 16#8205;   // Error: wrong length for write data record / Fehler: IO-Link-Master hat Fehlercode zurückgegeben, siehe "Diagnose"
      ERR_IO_LINK : Word := 16#8401;   // Error: IO-Link master returned error code, see "diagnostics" / Fehler: Gelesener Datensatz stimmt nicht mit Anfrage überein
      ERR_INCONSISTENT_DATA : Word := 16#8402;   // Error: Read data record doesn't match request / Fehler: Zeitüberschreitung bei Anforderung
      ERR_REQUEST_TIMEOUT : Word := 16#8403;   // Error: Request timed out / Fehler: Aufgrund eines undefinierten Zustands in der Zustandsmaschine
      ERR_UNDEFINED_STATE : Word := 16#8600;   // Error: due to an undefined state in state machine / Fehler: Aufgrund eines undefinierten Zustands in der Zustandsmaschine
      ERR_WRREC : Word := 16#8601;   // Error: WRREC encountered an error, see "diagnostics" / Fehler: WRREC hat einen Fehler festgestellt, siehe "Diagnose"
      ERR_RDREC : Word := 16#8602;   // Error: RDREC encountered an error, see "diagnostics" / Fehler: RDREC hat einen Fehler festgestellt, siehe "Diagnose"
      STATUS_MASK : DWord := 16#00FF_FF00;   // Mask to filter error codes / Maske zum Filtern von Fehlercodes
      STATUS_RESOURCE_BUSY : DWord := 16#0080_C200;   // Status from WRREC/RDREC: Resource is busy / Status von WRREC/RDREC: Ressource ist beschäftigt
      INDEX_CAP_IOLINK : Word := 16#B000;   // Index of the data record for IOLM_Info. Only IO-Link-Masters with CAP=16#B000 support this call. / Index des Datensatzes für IOLM_Info. Nur IO-Link-Master mit CAP=16#B000 unterstützen diesen Aufruf.
      CAP_LEGACY : Word := 16#00E3;   // Siemens (old) Standard CAP: 227 / Siemens (alt) Standard CAP: 227
      CAP_STANDARD : Word := 16#B400;   // IO-Link Standard CAP: 16#B400 / IO-Link-Standard-CAP: 16#B400
      STATUS_RDREC_VALID : Byte := 16#00;   // Status Code of RDREC in cased of no error occurs
      BITMASK_ERR_RDREC_B3 : Byte := 16#DE;   // Status Code of RDREC in case of an error when reading a data record
      BITMASK_ERR_RDREC_B2 : Byte := 16#80;   // Status Code of RDREC in case of an error when reading a data record - Error according to IEC 61158-6
      BITMASK_ERR_RDREC_B1 : Byte := 16#B0;   // Status Code of RDREC in case of an error when reading a data record - invalid index (cap)
   END_VAR
BEGIN
   REGION BLOCK INFO HEADER
       //===============================================================================
       // Siemens / (c)Copyright 2023
       //-------------------------------------------------------------------------------
       // Title:            LIOLink_Device
       // Function:         Acyclically reads or writes data records from and to IO-Link devices
       // Library:          LIOLink
       // Author:           Siemens Industry Online Support
       // Tested with:      CPU 1513-1 PN FW 2.8
       // Engineering:      TIA Portal V16
       // Restrictions:     S7-1200/1500
       // Requirements:     --
       //-------------------------------------------------------------------------------
       // Change log table:
       // Version  | Date       | Expert in charge       | Changes applied
       //----------|------------|------------------------|------------------------------
       // 02.00.00 | 30.09.2013 | Online Support         | First release for TIA Portal V12 SP1 as IO_LINK_CALL
       // 02.01.00 | 14.03.2014 | Online Support         | Upgrade to TIA Portal V13
       //                                                | Upgrade of system function 'WRREC' from V1.0 to V1.1
       // 03.00.00 | 28.02.2015 | SUP Applications       | Upgrade to TIA Portal V13 SP1
       //                                                | Renamed FB to IO_LINK_DEVICE 
       // 03.01.00 | 15.09.2015 | SUP Applications       | Change of #IOL_INDEX AND #Port lower boundry to 0 and improved behaviour when called in cyclic OBs with > 100 ms
       // 04.00.00 | 01.09.2020 | Online Support         | Implemented Programming styleguide for S7-1200/1500 and PLCopen
       //                                                | Renamed FB to LIOLink_Device 
       // 05.00.00 | 28.02.2023 | SUP SPH                | Added Polling Time as predefined input
       //                                                | #record is changed to a variable array (Array[*])
       //                                                | Changed CAP as predefined variable, added functionality to automatically find CAP of IO-Link-Masters from SIEMENS                                               
       //===============================================================================
   END_REGION

   REGION TRIGGERING
       #tempExecute := #execute; // Work with temporary value / create process image

       IF (#tempExecute = TRUE) AND (#statExecuteOld = FALSE) // Check if FB is triggered
           AND (#statStatus = #STATUS_NO_CALL)
       THEN
           REGION Initialize data
               // First call; initialize FB
               #statDone := FALSE;
               #statBusy := TRUE;
               #statError := FALSE;
               #statStatus := #STATUS_FIRST_CALL;
               #statSubfunctionStatus := #SUB_STATUS_NO_ERROR;
               #statFBErrorState := 0;
               #diagnostics := #statEmptyDiagnostics;
               #readLen := 0;

               // Initialize data area
               #statRead.header."call"."port" := 16#0;
               #statRead.header.iolHeader.indexLowByte := 16#0;
               #statRead.header.iolHeader.indexHighByte := 16#0;
               #statRead.header.iolHeader.subindex := 16#0;
               #tempIndexCounter := 0; // initialize loop counter      
               FOR #tempIndexCounter := 0 TO #UPPER_LIMIT DO
                   #statWrite.data[#tempIndexCounter] := 16#0;
                   #statRead.data[#tempIndexCounter] := 16#0;
               END_FOR;
           END_REGION

           REGION Save inputs
               // Copy input variables to temporary variables
               #tempHwID := #hwID;
               #statReadWrite := #readWrite;
               #statTimeout := #timeout;
               #statPollingPeriod := #pollingPeriod;
               #tempPort := #port;
               #tempIndex := #index;
               #tempSubindex := #subindex;
           END_REGION

           REGION Build header
               // setup call header
               #statWrite.header."call"."port" := INT_TO_BYTE(#tempPort);

               // setup IOL header 
               #statWrite.header.iolHeader.indexLowByte := INT_TO_BYTE(#tempIndex);
               #statWrite.header.iolHeader.indexHighByte := INT_TO_BYTE(SHR(IN := #tempIndex, N := 8));
               #statWrite.header.iolHeader.subindex := INT_TO_BYTE(#tempSubindex);

               // BODY (data max. 232 Byte, Array 0..231 of Byte) 
               IF #statReadWrite = #MODE_WRITE THEN // Write data record requested, copy data from "record"
                   #statWrite.header.iolHeader.control := #CONTROL_WRITE;
                   #statLen := INT_TO_UINT(#writeLen) + #LEN_HEADER; // data length header + data = IO-Link write data record
                   // copy "record" to working area
                   FOR #tempIndexCounter := 0 TO #writeLen - 1 DO
                       #statWrite.data[#tempIndexCounter] := #record[#tempIndexCounter];
                   END_FOR;
               ELSE // Read data record requested
                   // Empty record array
                   FILL_BLK(IN := 16#0,
                            COUNT := #MAX_DATA,
                            OUT => #record[0]);

                   #statWrite.header.iolHeader.control := #CONTROL_READ;
                   #statLen := #LEN_HEADER; // data length only header = IO-Link read data record
               END_IF;
           END_REGION

           REGION Check parameters
               // Check parameters
               IF (#tempPort < 0) OR (#tempPort > #MAX_PORT) THEN
                   #statStatus := #ERR_WRONG_PORT;
               ELSIF (#tempIndex < 0) OR (#tempIndex > #MAX_INDEX AND #tempIndex <> #INDEX_PORT_FUNC) THEN
                   #statStatus := #ERR_WRONG_INDEX;
               ELSIF (#tempSubindex < 0) OR (#tempSubindex > #MAX_SUBINDEX) THEN
                   #statStatus := #ERR_WRONG_SUBINDEX;
               ELSIF #statReadWrite = #MODE_WRITE AND (#writeLen < 1 OR #writeLen > #MAX_DATA) THEN
                   #statStatus := #ERR_WRONG_LENGTH;
               END_IF;
               //save the hwID from the previous execute
               #statHwIDprevious := #statHwID;

               IF #statStatus = #STATUS_FIRST_CALL THEN // Parameters OK
                   IF #cap <> 0 THEN
                       #statCap := INT_TO_UINT(#cap);
                       #statFBState := #FB_STATE_WRITE;
                   ELSIF (#statCap <> WORD_TO_UINT(#CAP_STANDARD) AND #statCap <> WORD_TO_UINT(#CAP_LEGACY)) OR (#statHwIDprevious <> #tempHwID) THEN // check if new device is connected => hwID changed
                       #statFBState := #FB_STATE_READ_CAP;
                   ELSE
                       #statFBState := #FB_STATE_WRITE;
                   END_IF;
               END_IF;
               // save current hwID
               #statHwID := #tempHwID;
           END_REGION

       ELSIF (#statStatus = #STATUS_FIRST_CALL) THEN
           #statStatus := #STATUS_SUBSEQUENT_CALL;
       END_IF;

       // Edge detection 'execute' input
       #statExecuteOld := #tempExecute;
   END_REGION TRIGGERING

   REGION STATE_MACHINE
       CASE #statFBState OF
           #FB_STATE_NO_PROCESSING:
               REGION no processing
                   ; // No processing active
               END_REGION no processing    

           #FB_STATE_READ_CAP:
               REGION get cap
                   // To find out CAP of IO-Link Master, data record with Index 16#B000 is read. If this reading was successful
                   // then CAP is 16#B400 (based on IO-Link Standard). If the reading was not successful and the status of RDREC
                   // is 16#DE80_B0xx, then CAP is 16#00E3 (227, based on Siemens Old Standard for IO-Link Masters).

                   #instRdRec(RECORD := #statRead);

                   IF (#instRdRec.BUSY = FALSE) THEN
                       IF (#instRdRec.VALID = FALSE) AND (#instRdRec.ERROR = FALSE) THEN
                           IF #instRdRec.REQ = FALSE THEN
                               // call read record with Index 16#B000
                               #instRdRec.REQ := true;
                               #instRdRec.ID := #statHwID;
                               #instRdRec.INDEX := WORD_TO_UINT(#INDEX_CAP_IOLINK);
                               #instRdRec.MLEN := 0;
                               #statFBState := #FB_STATE_READ_CAP;
                           END_IF;
                       ELSIF #instRdRec.VALID = TRUE THEN
                           #instRdRec.REQ := FALSE;
                           // if status of RDREC is valid then CAP is 16#B400 (CAP_STANDARD)
                           IF #instRdRec.STATUS.%B3 = #STATUS_RDREC_VALID THEN
                               #statCap := WORD_TO_UINT(#CAP_STANDARD);
                           END_IF;
                           #statFBState := #FB_STATE_WRITE;
                       ELSE
                           // if RDREC is in error state and Status is 16#DE80_B0xx then CAP is 227 (CAP_Legacy)
                           IF (#instRdRec.STATUS.%B3 = #BITMASK_ERR_RDREC_B3) AND (#instRdRec.STATUS.%B2 = #BITMASK_ERR_RDREC_B2) AND (#instRdRec.STATUS.%B1 = #BITMASK_ERR_RDREC_B1) THEN
                               #statCap := WORD_TO_UINT(#CAP_LEGACY);
                               #statFBState := #FB_STATE_WRITE;
                           ELSE
                               #statStatus := #ERR_RDREC;
                               #statSubfunctionStatus := #instRdRec.STATUS;
                               #statCap := 0; //clear CAP if an error occurs
                           END_IF;
                       END_IF;
                   ELSE
                       #instRdRec.REQ := FALSE;
                       IF #instRdRec.ERROR = TRUE THEN
                           #statStatus := #ERR_RDREC;
                           #statSubfunctionStatus := #instRdRec.STATUS;
                           #statCap := 0; //clear CAP if an error occurs
                       END_IF;
                   END_IF;

                   #instRdRec(RECORD := #statRead);
               END_REGION

           #FB_STATE_WRITE:
               REGION write
                   // To read data records, the IO-Link master modules needs to know which port is required. Therefore it is necessary
                   // to send at first a request via write data record (header, 8 byte). As response the IO-Link master module will 
                   // send the required data record.

                   #instWrRec(REQ := TRUE,
                              ID := #statHwID,
                              INDEX := #statCap,
                              LEN := #statLen,
                              RECORD := #statWrite);

                   IF #instWrRec.ERROR THEN
                       IF (#instWrRec.STATUS AND #STATUS_MASK) = #STATUS_RESOURCE_BUSY THEN
                           #instWrRec(REQ := FALSE); // Reset requeset
                       ELSE
                           #statStatus := #ERR_WRREC;
                           #statSubfunctionStatus := #instWrRec.STATUS;
                           #statFBErrorState := #statFBState;
                       END_IF;
                   ELSIF #instWrRec.DONE = TRUE THEN
                       #instWrRec(REQ := FALSE); // Reset requeset

                       #statFBState := #FB_STATE_POLL;
                   END_IF;
               END_REGION write

           #FB_STATE_POLL: // wait and poll for response
               REGION poll
                   #instPoll(IN := TRUE,
                             PT := #statPollingPeriod);

                   // read data record on falling edge
                   #instRdRec(REQ := NOT #instPoll.Q,
                              ID := #statHwID,
                              INDEX := #statCap,
                              MLEN := 0, // read all data available,
                              RECORD := #statRead);

                   IF #instRdRec.ERROR = TRUE THEN
                       IF (#instRdRec.STATUS AND #STATUS_MASK) = #STATUS_RESOURCE_BUSY THEN
                           // Reset requests and try again
                           #instPoll(IN := FALSE,
                                     PT := #statPollingPeriod);

                           #instRdRec(REQ := FALSE,
                                      RECORD := #statRead);
                       ELSE
                           #statStatus := #ERR_RDREC;
                           #statSubfunctionStatus := #instRdRec.STATUS;
                           #statFBErrorState := #statFBState;
                       END_IF;
                   ELSIF #instRdRec.VALID THEN
                       IF // check the response wether it matches the request (compare PORT, INDEX and SUBINDEX)
                           (#statWrite.header."call"."port" <> #statRead.header."call"."port")
                           OR (#statWrite.header.iolHeader.indexHighByte <> #statRead.header.iolHeader.indexHighByte)
                           OR (#statWrite.header.iolHeader.indexLowByte <> #statRead.header.iolHeader.indexLowByte)
                           OR (#statWrite.header.iolHeader.subindex <> #statRead.header.iolHeader.subindex)
                       THEN // read data record doesn't match the request
                           #statStatus := #ERR_INCONSISTENT_DATA;  // output status no consistent data
                       ELSIF #statRead.header.iolHeader.control = B#16#80 THEN // check the response for IO-Link errors
                           // State 0x80 = IOL_CALL_RES PDU shows IO-Link error detect
                           #statStatus := #ERR_IO_LINK;
                           #statSubfunctionStatus.%B3 := #statRead.data[0]; // IO-Link master error code
                           #statSubfunctionStatus.%B2 := #statRead.data[1]; // IO-Link master error code
                           #statSubfunctionStatus.%B1 := #statRead.data[2]; // ISDU error code
                           #statSubfunctionStatus.%B0 := #statRead.data[3]; // ISDU additional code
                           #statFBErrorState := #statFBState;
                       ELSE // read data is valid
                           IF #statReadWrite = #MODE_READ THEN
                               #readLen := UINT_TO_INT(#instRdRec.LEN - #LEN_HEADER);
                               // only data will be output
                               FOR #tempIndexCounter := 0 TO UINT_TO_INT(#instRdRec.LEN - #LEN_HEADER - 1) DO
                                   #record[#tempIndexCounter] := #statRead.data[#tempIndexCounter];
                               END_FOR;
                           END_IF;

                           // Reset requests
                           #instRdRec(REQ := FALSE,
                                      RECORD := #statRead);

                           #instPoll(IN := FALSE,
                                     PT := #statPollingPeriod);

                           #statStatus := #STATUS_EXECUTION_FINISHED;  // request finished
                       END_IF;
                   END_IF;
               END_REGION poll

           ELSE // Undefined state in state machine reached
               REGION undefined state
                   #statStatus := #ERR_UNDEFINED_STATE;
               END_REGION undefined state no relevant case, ready for new request
       END_CASE;
   END_REGION

   REGION MONITORING
       #instMonitor(IN := #statBusy,
                    PT := #statTimeout);

       IF #instMonitor.Q THEN
           #statStatus := #ERR_REQUEST_TIMEOUT; // request time out
       END_IF;
   END_REGION

   REGION OUTPUTS
       // Write outputs
       IF (#statStatus = #STATUS_EXECUTION_FINISHED) AND (#statDone = FALSE) THEN // Execution finished without errors, available only for one cycle
           REGION execution finished
               #statDone := TRUE;
               #statBusy := FALSE;
               #statError := FALSE;
               // execution aborted --> set state no processing
               #statFBState := #FB_STATE_NO_PROCESSING;
           END_REGION execution finished

       ELSIF (#statStatus.%X15 = TRUE) AND (#statError = FALSE) THEN // Error occurred (#statStatus is 16#8000 to 16#FFFF), Error status is true only for one cycle (the second last cycle)
           REGION error occured
               #statDone := FALSE;
               #statBusy := FALSE;
               #statError := TRUE;
               #statCap := 0; //Reset statcap, if error occurs, get cap has to be performed again
               // Write diagnostics
               #diagnostics.status := #statStatus;
               #diagnostics.subfunctionStatus := #statSubfunctionStatus;
               #diagnostics.stateNumber := #statFBErrorState;
               // Call instructions with FALSE to be ready for next job
               #instWrRec(REQ := FALSE);

               #instRdRec(REQ := FALSE,
                          RECORD := #statRead);

               #instPoll(IN := FALSE,
                         PT := #statPollingPeriod);

               // execution aborted --> set state no processing
               #statFBState := #FB_STATE_NO_PROCESSING;
           END_REGION error occured

       ELSIF (#tempExecute = FALSE) AND ((#statDone = TRUE) OR (#statError = TRUE)) THEN // Reset outputs, Last cycle
           REGION execute reset
               #statDone := FALSE;
               #statBusy := FALSE;
               #statError := FALSE;
               #statStatus := #STATUS_NO_CALL;
               #readLen := 0;
           END_REGION execute reset
       END_IF;

       REGION write static values to outputs
           #done := #statDone;
           #busy := #statBusy;
           #error := #statError;
           #status := #statStatus;
           //ENO := NOT #statError;
       END_REGION write static values to outputs
   END_REGION OUTPUTS
END_FUNCTION_BLOCK

// folder: LIOLink/S7-1200/1500/Device-specific blocks/SIMATIC RF200

FUNCTION_BLOCK "LIOLink_RF200_ReadTag"   // FB4, SCL
TITLE = LIOLink_RF200_ReadTag
{ S7_Optimized_Access := 'TRUE' }
AUTHOR : SIOS
FAMILY : LIOLink
VERSION : 3.0
// Reads tags from SIMATIC RF200 readers via IO-Link
   VAR_INPUT
      execute : Bool;   // Request job (on rising edge)
      addrTag : Word;   // Start address of data on tag
      length : Word;   // Length of data to be read
      hwID : HW_SUBMODULE;   // Logic IO address of the IO-Link Master
      portAddr : Int;   // Start address of port
      "version" : USInt := 11;   // IO-Link version of the reader; 11: IO-Link V1.1, 10: IO-Link V1.0
   END_VAR
   VAR_OUTPUT
      done : Bool;   // FALSE: data invalid, TRUE: data valid
      busy : Bool;   // FALSE: no job, TRUE: job in progress
      error : Bool;   // FALSE: no error, TRUE: error
      status : DWord;   // Error status
      presence : Bool;   // TRUE: Transponder on field
   END_VAR
   VAR_IN_OUT
      identData : Variant;   // Received tag identification data
   END_VAR
   VAR
      statPae : Array[0..#UPPER_BOUND_NETTO_IO_FIELD] of Byte;   // Partly recived identification data vie Process image
      statStatusByte : Byte;   // RF200 Tag reader status byte
      statPresence : Bool;   // TRUE: Transponder on field
      statState : Int;   // Main State Machine Index
      statAddr : Word;   // Start address of data on tag
      statOffset : Int;   // Buffer offset
      statExecuteReq : Bool;   // Execute function memory
      statLength : DInt;   // Length of read data
      statDat : Array[0..#UPPER_BOUND_IO_FIELD] of Byte;   // Data to Send
      statRecDat : Array[0..#UPPER_BOUND_IO_FIELD] of Byte;   // Data Received
      statAddrOffset : Int;   // Start adress of port
      statPresenceFF : Bool;   // TRUE: Transponder on field
      instTonrTime : TONR_TIME;   // Tag has left antenna field detection timer
      statTimerIn : Bool;   // Tag has left antenna field detection timer - Start Tag
      statTimerR : Bool;   // Tag has left antenna field detection timer - Reset Tag
      statTimerPt : Time := T#5S;   // Tag has left antenna field detection timer - Detection time
      statReadData : Array[0..#UPPER_BOUND_MAX_DATA_FIELD] of Byte;   // Received tag identification data
      statCountCopyPae : DInt;   // Length of current next data part in process image
      statBusy : Bool;   // TRUE: FB is not finished and new output values can be expected
      statDone : Bool;   // TRUE: Commanded functionality has been completed successfully
      statError : Bool;   // TRUE: Commanded functionality has been canceled with error
      statReturnMoveBlkVar : Int;   // Return Value PAE copy function
      statDiffToIOsizeNetto : Int;   // Difference between requested length and PAE
      instSetIoPart : SETIO_PART;   // Instance for PIQ writing
      statIoPartError : Bool;   // TRUE: data in process image is invalid
      statIoPartStatus : DWord;   // Status for IO access
      instGetIoPart : GETIO_PART;   // Instance for PII reading
      statIOsize : USInt;   // Size of the IO-Link Master PII
      statIOsizeNetto : USInt;   // Size of the IO-Link Master PAE without header
   END_VAR
   VAR_TEMP
      tempStatus : DWord;   // Auxiliary tag for status output
   END_VAR
   VAR CONSTANT
      IOL_V10 : USInt := 10;   // Identifier IO-Link version 1.0
      IOL_V11 : USInt := 11;   // Identifier IO-Link version 1.1
      LEN_DATA_V10 : USInt := 8;   // Length of user data for IO-Link version 1.0
      LEN_DATA_V11 : USInt := 32;   // Length of user data for IO-Link version 1.1
      UPPER_BOUND_IO_FIELD : USInt := 31;   // Upper bound of Input and Output fields
      UPPER_BOUND_NETTO_IO_FIELD : USInt := 27;   // Upper bound of Input and Output fields without header
      UPPER_BOUND_MAX_DATA_FIELD : UInt := 1999;   // Upper bound of the data field of a RFID Tag
      DATA_HEADER_SIZE : USInt := 4;   // IO-Link Header Size for version 1.0 and 1.1
      CMD_READ : Byte := 16#02;   // Command to read data
      CMD_RESET : Byte := 16#00;   // Command to reset
      MIN_LENGTH_V10 : Word := 16#0004;   // Minimal Lenght of requested tag information
      MIN_LENGTH_V11 : Word := 16#001C;   // Minimal Lenght of requested tag information
      STATUS_ERROR_IDENT_BLOCK : Word := 16#0001;   // Error Identification for block internal faults
      STATUS_ERROR_IDENT_RFID : Word := 16#0011;   // Error Identification for RFID reader faults
      STATUS_NO_JOB : Word := 16#0000;   // No job requested
      STATUS_ERROR_TAG_HAS_LEFT : Word := 16#8101;   // Error - the RFID tag has left the reader
      STATUS_ERROR_STILL_ACTIVE : Word := 16#8102;   // Error - block still busy, no further request possible
      STATUS_ERROR_LENGTH : Word := 16#8104;   // Error - requested length is less than 0
      STATE_IDLE : Int := 0;   // State Machine - Idle State
      STATE_READ : Int := 2;   // State Machine - Read Tag
      STATE_TELEGRAM : Int := 1;   // State Machine - Prepare telegram
      STATE_ERROR : Int := 3;   // State Machine - Error State
      DETECTION_TIME_TAG_OFF_FIELD : Time := T#5S;   // Tag has left antenna field detection time
      INDEX_CMD : USInt := 0;   // Index in DataField - Command
      INDEX_RFID_ERROR : USInt := 1;   // Index in DataField - Error
      INDEX_ADDR_HIGH : USInt := 2;   // Index in DataField - Address High Byte
      INDEX_ADDR_LOW : USInt := 3;   // Index in DataField - Address Low Byte
      INDEX_SOURCE_DATA : DInt := 4;   // Index in Data Field - Start of netto Data
   END_VAR
BEGIN
   REGION BLOCK INFO HEADER
       //===============================================================================
       // Siemens / (c)Copyright 2022
       //-------------------------------------------------------------------------------
       // Title:            LIOLink_RF200_ReadTag
       // Function:         Reads tags from SIMATIC RF200 readers via IO-Link
       // Library:          LIOLink
       // Author:           Siemens Industry Online Support
       // Tested with:      CPU 1513-1 PN FW 2.8
       // Engineering:      TIA Portal V16
       // Restrictions:     --
       // Requirements:     --
       //-------------------------------------------------------------------------------
       // Change log table:
       // Version  | Date       | Expert in charge       | Changes applied
       //----------|------------|------------------------|------------------------------
       // 01.00.00 | 01.07.2013 | Online Support         | First release
       // 01.01.00 | 01.12.2016 | Online Support         | Upgraded to TIA Portal V14
       // 02.00.00 | 01.09.2017 | Online Support         | Upgraded to TIA Portal V14 SP1
       //                                                | Implemented Programming styleguide
       //                                                | Added support for IO-Link V1.1 readers
       // 02.01.00 | 01.12.2017 | Online Support         | Bug fixes and performance improvements
       // 02.02.00 | 01.03.2020 | Online Support         | Upgraded to TIA Portal V16
       // 02.03.00 | 22.09.2020 | Online Support         | Integrated FB into LIOLink library
       //                                                | Renamed FB to LIOLink_RF200_ReadTag
       //                                                | Combined FBs for IO-Link V1.0 and V1.1
       //                                                | Minor bug fixes
       // 02.04.00 | 29.06.2022 | Online Support         | Minor bug fixes     
       // 02.05.00 | 30.09.2022 | SUP SPH                | Optimization     
       //===============================================================================
   END_REGION

   REGION Check version
       //determine IO-Link reader version (1.0/1.1) to set offsets
       IF #version = #IOL_V11 THEN
           #statIOsize := #LEN_DATA_V11;
           #statIOsizeNetto := #LEN_DATA_V11 - #DATA_HEADER_SIZE;
       ELSE
           #statIOsize := #LEN_DATA_V10;
           #statIOsizeNetto := #LEN_DATA_V10 - #DATA_HEADER_SIZE;
       END_IF;
   END_REGION

   REGION Get PII
       #statAddrOffset := #portAddr;   //start adress of port

       // Read PII
       #instGetIoPart(ID := #hwID,
                      OFFSET := #statAddrOffset,
                      LEN := #statIOsize,
                      STATUS => #statIoPartStatus,
                      ERROR => #statIoPartError,
                      INPUTS := #statRecDat);

       #statStatusByte := #statRecDat[0];    //Status Byte
       #statPresence := #statStatusByte.%X5;   //Presence bit. Transponder on field
   END_REGION

   REGION Check execute
       REGION Idle
           IF NOT #execute THEN
               #statDone := false;
               #statBusy := false;
               #statError := false;
               #tempStatus := #STATUS_NO_JOB;
           END_IF;
       END_REGION

       REGION Job requested
           //Positive edge for reading of data
           IF #execute AND #execute <> #statExecuteReq THEN
               IF NOT #statBusy THEN
                   #statAddr := #addrTag;    //Transpoder Address
                   #statDiffToIOsizeNetto := WORD_TO_INT(#length) MOD #statIOsizeNetto;
                   #statLength := WORD_TO_DINT(#length);   //Length of read Dat
                   #statBusy := TRUE;
                   #statDone := FALSE;
                   #statError := FALSE;
                   #tempStatus := #STATUS_NO_JOB;
                   #statOffset := 0;   //offset of puffer must be reseted
                   #statState := #STATE_READ;    //next step >> send read command
                   #statCountCopyPae := 0;
                   FILL_BLK(IN := 0,    //Reset read buffer
                            COUNT := CountOfElements(#identData),
                            OUT => #statReadData[0]);
               ELSE
                   #tempStatus.%W0 := #STATUS_ERROR_STILL_ACTIVE;                       //block is still active
                   #tempStatus.%W1 := #STATUS_ERROR_IDENT_BLOCK;                        //Error identifier for block errors
                   #statState := #STATE_ERROR;
               END_IF;
               IF #length < 0 OR (#length < #MIN_LENGTH_V11 AND #version = #IOL_V11) OR (#length < #MIN_LENGTH_V10 AND #version = #IOL_V10) THEN
                   #tempStatus.%W0 := #STATUS_ERROR_LENGTH;                             //length too short
                   #tempStatus.%W1 := #STATUS_ERROR_IDENT_BLOCK;                        //identifier rfid errors
                   #statState := #STATE_ERROR;
               END_IF;
           END_IF;
       END_REGION
       #statExecuteReq := #execute;
   END_REGION

   REGION Tag presence detection
       IF NOT #statPresence AND #statPresence <> #statPresenceFF THEN   //the tag has left the antenna  field
           IF NOT #statDone THEN
               #statTimerIn := true;   //wait 5 sec
               #statTimerR := false;
           END_IF;
       END_IF;
       #statPresenceFF := #statPresence;
       IF #statPresence THEN
           #statTimerR := true;
           #statTimerIn := false;
       END_IF;
   END_REGION

   REGION State machine
       CASE #statState OF
           #STATE_IDLE:
               #statBusy := false;
               #statTimerIn := false;

           #STATE_READ:
               IF #statLength > 0 THEN
                   #statDat[#INDEX_CMD] := #CMD_READ;    //Set read command
                   #statDat[#INDEX_ADDR_HIGH] := #statAddr.%B1;    //Adr-H
                   #statDat[#INDEX_ADDR_LOW] := #statAddr.%B0;   //Adr-L
               END_IF;

               IF NOT #statIoPartError THEN
                   #statState := #STATE_TELEGRAM;    //Telegram: Edit the read data
               END_IF;

           #STATE_TELEGRAM:
               IF #statLength > 0 THEN   //Only when length of data>0 can continue  
                   IF #statStatusByte.%X6 THEN   //IF RFID error has occured
                       #tempStatus.%W0 := #statRecDat[#INDEX_RFID_ERROR];    //error_RFID
                       #tempStatus.%W1 := #STATUS_ERROR_IDENT_RFID;    //Error identifier for RFID errors
                       #statState := #STATE_ERROR;
                   END_IF;

                   //-------------------------- read command is ready------------------------------------------------//
                   IF #statStatusByte.%X7 AND #statStatusByte.%X1 THEN
                       IF #statRecDat[#INDEX_ADDR_HIGH] = #statAddr.%B1
                           AND #statRecDat[#INDEX_ADDR_LOW] = #statAddr.%B0
                       THEN //received ADR must be ==sent ADR
                           #statReturnMoveBlkVar := MOVE_BLK_VARIANT(SRC := #statRecDat,
                                                                     COUNT := #statIOsizeNetto,
                                                                     SRC_INDEX := #INDEX_SOURCE_DATA,
                                                                     DEST_INDEX := 0,
                                                                     DEST => #statPae);

                           IF NOT #statIoPartError THEN
                               IF #statCountCopyPae = 0 THEN    //copy the #statIOsizeNet Bytes in 
                                   IF #statLength >= #statIOsizeNetto THEN
                                       IF #statLength <> WORD_TO_DINT(#length) THEN
                                           #statAddr := INT_TO_WORD(WORD_TO_INT(#statAddr) + #statIOsizeNetto);
                                       END_IF;
                                       #statState := #STATE_READ;
                                       #statCountCopyPae := #statIOsizeNetto;
                                   ELSE
                                       IF #statStatusByte.%X7 AND NOT #statStatusByte.%X6 THEN
                                           IF #statDiffToIOsizeNetto <> 0 THEN
                                               #statCountCopyPae := #statDiffToIOsizeNetto;
                                               #statAddr := INT_TO_WORD(WORD_TO_INT(#statAddr) + #statIOsizeNetto);
                                               #statState := #STATE_READ;
                                           ELSE
                                               #statCountCopyPae := #statIOsizeNetto;
                                           END_IF;
                                       ELSE
                                           #statState := #STATE_IDLE;
                                       END_IF;
                                   END_IF;
                               ELSE
                                   #statReturnMoveBlkVar := MOVE_BLK_VARIANT(SRC := #statPae,
                                                                             COUNT := DINT_TO_UDINT(#statCountCopyPae),
                                                                             SRC_INDEX := 0,
                                                                             DEST_INDEX := #statOffset,
                                                                             DEST => #statReadData);
                                   IF #statReturnMoveBlkVar = 0 THEN
                                       #statCountCopyPae := 0;
                                       #statOffset := #statOffset + #statIOsizeNetto;
                                       #statLength := #statLength - #statIOsizeNetto;
                                   END_IF;
                               END_IF;
                           ELSE
                               #tempStatus.%W0 := DWORD_TO_WORD(#statIoPartStatus);    //Error has to BLKMOV occured
                               #tempStatus.%W1 := #STATUS_ERROR_IDENT_BLOCK;   //functions-Error identifier
                               #statState := #STATE_ERROR;
                           END_IF;
                       END_IF;
                   END_IF;
                   #instSetIoPart(ID := #hwID,
                                  OFFSET := #statAddrOffset,
                                  LEN := #statIOsize,
                                  STATUS => #statIoPartStatus,
                                  ERROR => #statIoPartError,
                                  OUTPUTS := #statDat);

                   IF #statIoPartError THEN
                       #tempStatus.%W0 := DWORD_TO_WORD(#statIoPartStatus);    //Error has to BLKMOV occured
                       #tempStatus.%W1 := #STATUS_ERROR_IDENT_BLOCK;   //functions-Error identifier
                       #statState := #STATE_ERROR;
                   END_IF;

               ELSE
                   VariantPut(SRC := #statReadData,
                              DST := #identData);
                   #statState := #STATE_IDLE;
                   #statBusy := false;
                   #statDone := true;

                   //Reset read command
                   #statDat[#INDEX_CMD] := #CMD_RESET;

                   #instSetIoPart(ID := #hwID,
                                  OFFSET := #statAddrOffset,
                                  LEN := #statIOsize,
                                  STATUS => #statIoPartStatus,
                                  ERROR => #statIoPartError,
                                  OUTPUTS := #statDat);
               END_IF;

           #STATE_ERROR:
               #statBusy := false;
               #statDone := false;
               #statError := true;
               #statTimerIn := false;
               #statTimerR := true;
               #statState := #STATE_IDLE;

               //Reset read command
               #statDat[#INDEX_CMD] := #CMD_RESET;

               #instSetIoPart(ID := #hwID,
                              OFFSET := #statAddrOffset,
                              LEN := #statIOsize,
                              STATUS => #statIoPartStatus,
                              ERROR => #statIoPartError,
                              OUTPUTS := #statDat);
           ELSE
               #statState := #STATE_IDLE;
       END_CASE;
   END_REGION

   REGION Detection timer
       #instTonrTime(IN := #statTimerIn,   //this timer will start, if the tag has left the antenna field
                     R := #statTimerR,
                     PT := #statTimerPt);
       IF #instTonrTime.Q THEN   //error has occured. No tag on field during the 5 sec.
           #tempStatus.%W0 := #STATUS_ERROR_TAG_HAS_LEFT;    //tag has left the field
           #tempStatus.%W1 := #STATUS_ERROR_IDENT_BLOCK;   //identifier rfid errors
           #statState := #STATE_ERROR;
       END_IF;
   END_REGION

   REGION Update output interface 
       #done := #statDone;
       #busy := #statBusy;
       #error := #statError;
       #status := #tempStatus;
       #presence := #statPresence;
   END_REGION
END_FUNCTION_BLOCK

FUNCTION_BLOCK "LIOLink_RF200_SwitchAntenna"   // FB5, SCL
TITLE = LRfidIOL_ANT
{ S7_Optimized_Access := 'TRUE' }
AUTHOR : SIOS
FAMILY : LIOLink
VERSION : 3.1
// Set Antenna
// IO-Link V1.1
   VAR_INPUT
      execute : Bool;   // Execute function
      antennaState : Bool;   // TRUE: activate antenna, FALSE: deactivate antenna
      hwID : HW_SUBMODULE;   // Hardware identifier of IO-Link communication module
      portAddr : Int;   // Start address of port
      "version" : USInt := 11;   // IO-Link version of the reader; 11: IO-Link V1.1, 10: IO-Link V1.0
   END_VAR
   VAR_OUTPUT
      done : Bool;   // TRUE: Job done
      busy : Bool;   // TRUE: Job active
      error : Bool;   // TRUE: Error has occured
      status : DWord;   // Error status
      presence : Bool;   // TRUE: Transponder on field
   END_VAR
   VAR
      statExecuteReq : Bool;   // State of execute input of last cycle
      statAntStatus : Byte;   // Status Byte of antenna
      statState : UInt;   // Main State Machine Index
      statAnt : Array[0..#UPPER_BOUND_IO_FIELD] of Byte;   // Received buffer of Antenna data
      statSent : Array[0..#UPPER_BOUND_IO_FIELD] of Byte;   // Sent buffer for Antenna
      statPresence : Bool;   // Presence bit. Transponder on field
      statBusy : Bool;   // TRUE: Job active
      instSetIoPart : SETIO_PART;   // Instance for PIQ writing
      statIoPartError : Bool;   // TRUE: data in process image is invalid
      statIoPartStatus : DWord;   // Status for IO access
      instGetIoPart : GETIO_PART;   // Instance for PII reading
      statIOsize : Int;   // Size of the IO-Link Master PII
   END_VAR
   VAR_TEMP
      tempDone : Bool;   // Auxiliary tag for done output
      tempError : Bool;   // Auxiliary tag for error output
      tempStatus : DWord;   // Auxiliary tag for status output
   END_VAR
   VAR CONSTANT
      IOL_V10 : USInt := 10;   // Identifier IO-Link version 1.0
      IOL_V11 : USInt := 11;   // Identifier IO-Link version 1.1
      LEN_DATA_V10 : USInt := 8;   // Length of user data for IO-Link version 1.0
      LEN_DATA_V11 : USInt := 32;   // Length of user data for IO-Link version 1.1
      UPPER_BOUND_IO_FIELD : USInt := 31;   // Upper bound of Input and Output fields
      STATE_IDLE : UInt := 0;   // State Machine - Idle State
      STATE_ANTENNA_ON : UInt := 1;   // State Machine - Switch Antenna on
      STATE_ANTENNA_OFF : UInt := 2;   // State Machine - Switch Antenna off
      STATE_READY : UInt := 3;   // State Machine - Job done
      STATUS_ERROR_IDENT_BLOCK : Word := 16#0001;   // Error Identification for block internal faults
      STATUS_ERROR_IDENT_RFID : Word := 16#0011;   // Error Identification for RFID reader faults
      STATUS_NO_JOB : Word := 16#0000;   // No job requested
      STATUS_ERROR_TAG_HAS_LEFT : Word := 16#8101;   // Error - the RFID tag has left the reader
      STATUS_ERROR_STILL_ACTIVE : Word := 16#8102;   // Error - block still busy, no further request possible
      STATUS_ERROR_LENGTH : Word := 16#8104;   // Error - requested length is less than 0
      CMD_ANTENNA_ON : Byte := 16#00;   // Command to switsch antenna on
      CMD_ANTENNA_OFF : Byte := 16#10;   // Command to switsch antenna off
      INDEX_ANT_STATUS : USInt := 0;   // Index in Antenna DataField - Status
      INDEX_RFID_ERROR : USInt := 1;   // Index in Antenna DataField - Error
      INDEX_SEND_CMD : USInt := 0;   // Index in Send DataField - Command
   END_VAR
BEGIN
   REGION BLOCK INFO HEADER
       //===============================================================================
       // Siemens / (c)Copyright 2022
       //-------------------------------------------------------------------------------
       // Title:            LIOLink_RF200_SwitchAntenna
       // Function:         Switches the antenna of SIMATIC RF200 readers via IO-Link
       // Library:          LIOLink
       // Author:           Siemens Industry Online Support
       // Tested with:      CPU 1513-1 PN FW 2.8
       // Engineering:      TIA Portal V16
       // Restrictions:     --
       // Requirements:     --
       //-------------------------------------------------------------------------------
       // Change log table:
       // Version  | Date       | Expert in charge       | Changes applied
       //----------|------------|------------------------|------------------------------
       // 01.00.00 | 01.07.2013 | Online Support         | First release
       // 01.01.00 | 01.12.2016 | Online Support         | Upgrade to TIA Portal V14
       // 02.00.00 | 01.09.2017 | Online Support         | Upgrade to TIA Portal V14 SP1
       //                                                | Implementation of Programming styleguide
       //                                                | Added support for IO-Link V1.1 readers
       // 02.01.00 | 01.12.2017 | Online Support         | Bug fixes and performance improvements
       // 02.02.00 | 01.03.2020 | Online Support         | Upgrade to TIA Portal V16
       // 02.03.00 | 22.09.2020 | Online Support         | Integrated FB into LIOLink library
       //                                                | Renamed FB to LIOLink_RF200_SwitchAntenna
       //                                                | Combined FBs for IO-Link V1.0 and V1.1
       //                                                | Minor bug fixes
       // 02.04.00 | 04.10.2022 | SUP SPH                | Optimization
       //===============================================================================
   END_REGION

   REGION Check version
       IF #version = #IOL_V11 THEN                               //determine IO-Link reader version (1.0/1.1) to set offset
           #statIOsize := #LEN_DATA_V11;
       ELSE
           #statIOsize := #LEN_DATA_V10;
       END_IF;
   END_REGION

   REGION Get PII

